FUNCTION_BLOCK fbScheduler
VAR
	_Active : BOOL;
	_Now : TIMESTRUCT;
	NowTOD : TIME_OF_DAY;
	i : USINT;
	TimeDiff : DINT;
	ActiveRTrigger : R_TRIG;
END_VAR
VAR RETAIN
    _Enabled : BOOL := FALSE;
    _Config : stSchedulerConfig;
END_VAR
VAR CONSTANT
	EmptyTimeTrigger : TIME_OF_DAY := TOD#00:00;
	TriggerTimeTolerance : TIME := T#1M; 
END_VAR


_Active := FALSE;
NowTOD := SYSTEMTIME_TO_TOD(_Now);

// Sprawdz, czy trigger wlaczony
IF NOT _Enabled THEN 
  RETURN; 
END_IF;

// Sprawdz, czy aktualny miesiac
IF NOT _Config.Months[_Now.wMonth] THEN 
  RETURN; 
END_IF;

// Sprawdz, czy aktualny dzien
IF NOT _Config.WeekDays[_Now.wDayOfWeek + 1] THEN // (Now.wDayOfWeek 0 (Sunday) = CyclicTrigger.WeekDays[1])
  RETURN; 
END_IF;

// Sprawdz czasy
FOR i := 1 TO 6 DO
  IF _Config.Times[i] <> EmptyTimeTrigger THEN
	  TimeDiff := TOD_TO_DINT(NowTOD) - TOD_TO_DINT(_Config.Times[i]);	  
	  // Korekta przekroczenia doby (86 400 000 ms = 24h)
	IF TimeDiff > 43200000 THEN       // >12h różnicy → cofnij o dobę
		TimeDiff := TimeDiff - 86400000;
	ELSIF TimeDiff < -43200000 THEN   // <-12h różnicy → dodaj dobę
		TimeDiff := TimeDiff + 86400000;
	END_IF
	IF ABS(TimeDiff) <= TIME_TO_DINT(TriggerTimeTolerance) THEN  // ← TO BRAKOWAŁO
        _Active := TRUE;
        EXIT;  // Pierwsza zgodnosc wystarczy
    END_IF
  END_IF;
END_FOR;

ActiveRTrigger(CLK := _Active);

PROPERTY Enable : BOOL
GET
Enable := THIS^._Enabled;
END_GET
SET
THIS^._Enabled := Enable;
END_SET
END_PROPERTY

PROPERTY IsActive : BOOL
GET
IsActive := THIS^._Active;
END_GET
END_PROPERTY

METHOD SetConfig
VAR_INPUT
	Config : stSchedulerConfig;
END_VAR
THIS^._Config := Config;
END_METHOD

PROPERTY Triggered : BOOL
GET
Triggered := THIS^.ActiveRTrigger.Q;
END_GET
END_PROPERTY

METHOD UpdateTime
VAR_INPUT
	Now : TIMESTRUCT;
END_VAR
_Now := Now;
END_METHOD

END_FUNCTION_BLOCK

(* stored: Version 1.1.0.1
   POU fbScheduler: Id {e6beab7c-6878-4fdf-b4e1-89106bd737c9}, SpecialFunc None
   Property Enable: Id {2e980649-b9bf-4864-9037-87be4a693a3a}
   Get Get: Id {f622a717-b980-4bf5-8bc8-af059c50987c}
   Set Set: Id {f8d081ad-dbd1-4281-97d1-0f22ba6611a9}
   Property IsActive: Id {1670c2e2-c25a-4a5e-84dc-d3f2300321a8}
   Get Get: Id {62b511ae-b1df-442d-9bd8-f2eff94c4283}
   Method SetConfig: Id {1f07cda4-afa7-4310-8fba-eb5cd655d675}
   Property Triggered: Id {2975e954-9b3b-4e9b-b472-d35dfc8b1e42}
   Get Get: Id {1fa6a10c-de63-4b3a-a0b0-2bb8f0332aae}
   Method UpdateTime: Id {9c526424-860f-4349-8539-a9d423bc789c} *)
